(* IEC 61131-3 sources: JingjiangArm/moonboxpro_arm_8.4/Application/Application/任务列表/ExtTask/动作处理/涂布, 11 files *)

(* ---- StCoatingAxisInf.st ---- *)
(*@CES
Name=StCoatingAxisInf
Type=Gvl
TypeGuid=2db5746d-d284-4425-9f7f-2663a34b0ebc
Guid=2e9ecafb-d2f1-4b6b-83e3-f47895db637f
HasDeclaration=True
HasImplementation=False
*)
{DECLARATION}
TYPE StCoatingAxisInf :
STRUCT
(*涂布轴信息@2024.01.18.095207*)
	byCoatingAxisNum			: BYTE;(*涂布轴个数*)
	aiAxisIdList				: ARRAY [1..gc_byCoatingMaxSum_New]OF INT;(*轴idlist*)
	astStCoatingAxisParam		: ARRAY [1..gc_byCoatingMaxSum_New] OF StCoatingAxisParam;
END_STRUCT
END_TYPE

{IMPLEMENTATION}

(* ---- StCoatingAxisParam.st ---- *)
(*@CES
Name=StCoatingAxisParam
Type=Gvl
TypeGuid=2db5746d-d284-4425-9f7f-2663a34b0ebc
Guid=8a071cba-fd95-4a8c-93c6-fe3e9b0305b5
HasDeclaration=True
HasImplementation=False
*)
{DECLARATION}
{attribute 'pack_mode' := '1'}
TYPE StCoatingAxisParam :(*涂布轴参数@2024.01.18.093551*)
STRUCT
	iUnitId							:INT;(*轴id@默认-1*)
	xSwitchOn_CoatingPrn			:BOOL;(*涂布开关*)
	byAdjMode_CoatingPrn			:BYTE;(*涂布轴模式*)
	xReverseAdj_CoatingPrn			:BOOL;(*涂布轴调整取反*)
	rAI_CoatingPrn					:REAL;(*涂布轴模拟量*)
	rAI_med_CoatingPrn				:REAL;(*涂布轴中位值*)
	lrGirth_Using_CoatingPrn		:LREAL;(*涂布轴周长@界面输入*)
	iKp_CoatingPrn					:INT;(*涂布kp*)
	iKi_CoatingPrn					:INT;(*涂布ki*)
	iKd_CoatingPrn					:INT;(*涂布kd*)
	xFlag_PressDne					:BOOL;(*涂布轴合压*)

	rAI_CoatingHMI					:REAL;(*涂布模拟量显示*)
	lrGirth_CoatingPrn				:LREAL;(*涂布周长@用于运算pt*)
	lrVelocity_CoatingPrn			:LREAL;(*涂布速度*)
END_STRUCT
END_TYPE

{IMPLEMENTATION}

(* ---- KS_CoatingAxisParamDeal.st ---- *)
(*@CES
Name=KS_CoatingAxisParamDeal
Type=FunctionBlock
TypeGuid=6f9dac99-8de1-4efc-8465-68ac443b7d08
Guid=f4156371-7451-43fd-b965-d24d4d478a2f
HasDeclaration=True
HasImplementation=True
*)
{DECLARATION}
FUNCTION KS_CoatingAxisParamDeal : BOOL
VAR_INPUT
(*涂布轴参数处理*)
	i_byDealType:BYTE;(*处理方式@=1 初始化涂布轴参数
								@=2 从轴参数写入到涂布轴参数中#涂布控制输入变量
								@=3 涂布轴参数写入到轴参数中#涂布控制输出变量
								@=4 操作的轴参数值复位*)
	i_iAxisId:INT;
	i_xFlag_AxisPressDne:BOOL;(*轴的合压状态@经过延时后输出标志*)
	i_pstStCoatingAxisParam:POINTER TO StCoatingAxisParam;
	i_palrGirth_CoatingPrn:POINTER TO ARRAY [1..MAX_UNIT_NUM] OF LREAL;(*用于计算pt的周长值@未定义到轴参数中*)
	i_palrAI_CoatingHMI:POINTER TO ARRAY [1..MAX_UNIT_NUM] OF LREAL;(*界面显示的模拟量值@未定义到轴参数中*)
//2025.7.3.175755
	i_axSwitchOn_CoatingPrn: ARRAY [1..MAX_UNIT_NUM] OF BOOL;(*涂布开关*)
	i_abyAdjMode_CoatingPrn: ARRAY [1..MAX_UNIT_NUM] OF BYTE;(*涂布轴模式*)
	i_axReverseAdj_CoatingPrn: ARRAY [1..MAX_UNIT_NUM] OF BOOL;(*涂布轴调整取反*)
	i_alrAI_CoatingPrn: ARRAY [1..MAX_UNIT_NUM] OF LREAL;(*涂布模拟量*)
	i_alrAI_med_CoatingPrn: ARRAY [1..MAX_UNIT_NUM] OF LREAL;(*涂布中位值*)
	i_alrGirth_Using_CoatingPrn: ARRAY [1..MAX_UNIT_NUM] OF LREAL;(*涂布轴周长*)
	i_aiKp_CoatingPrn: ARRAY [1..MAX_UNIT_NUM] OF INT;(*涂布Kp*)
	i_aiKi_CoatingPrn: ARRAY [1..MAX_UNIT_NUM] OF INT;(*涂布Ki*)
	i_aiKd_CoatingPrn: ARRAY [1..MAX_UNIT_NUM] OF INT;(*涂布Kd*)
	i_palrVelocity_CoatingPrn:POINTER TO ARRAY [1..MAX_UNIT_NUM] OF LREAL;(*涂布轴速度*)
	i_alrGirth:ARRAY [1..MAX_UNIT_NUM] OF LREAL;(*当前轴周长*)
END_VAR
VAR
END_VAR

{IMPLEMENTATION}
CASE i_byDealType OF
	1:(*初始化涂布参数*)
		IF i_pstStCoatingAxisParam<>0 THEN
			SysMemSet(i_pstStCoatingAxisParam,0,SIZEOF(i_pstStCoatingAxisParam^));
			i_pstStCoatingAxisParam^.iUnitId:=-1;
		END_IF
	2:(*从轴参数写入到涂布轴参数中#涂布控制输入变量*)
		IF i_iAxisId>0 AND i_iAxisId<MAX_UNIT_NUM AND(*轴号合法*)

			i_pstStCoatingAxisParam<>0 THEN

			i_pstStCoatingAxisParam^.iUnitId						:= i_iAxisId;
			i_pstStCoatingAxisParam^.xSwitchOn_CoatingPrn			:= i_axSwitchOn_CoatingPrn[i_iAxisId];(*涂布开关*)
			i_pstStCoatingAxisParam^.byAdjMode_CoatingPrn			:= i_abyAdjMode_CoatingPrn[i_iAxisId];(*涂布轴模式*)
			i_pstStCoatingAxisParam^.xReverseAdj_CoatingPrn			:= i_axReverseAdj_CoatingPrn[i_iAxisId]	;(*涂布轴调整取反*)
			i_pstStCoatingAxisParam^.rAI_CoatingPrn					:= i_alrAI_CoatingPrn[i_iAxisId];(*涂布轴模拟量*)
			i_pstStCoatingAxisParam^.rAI_med_CoatingPrn				:= i_alrAI_med_CoatingPrn[i_iAxisId];(*涂布轴中位值*)
			i_pstStCoatingAxisParam^.lrGirth_Using_CoatingPrn		:= i_alrGirth_Using_CoatingPrn[i_iAxisId];(*涂布轴周长@界面输入*)
			i_pstStCoatingAxisParam^.iKp_CoatingPrn					:= i_aiKp_CoatingPrn[i_iAxisId]	;(*涂布kp*)
			i_pstStCoatingAxisParam^.iKi_CoatingPrn					:= i_aiKi_CoatingPrn[i_iAxisId];(*涂布ki*)
			i_pstStCoatingAxisParam^.iKd_CoatingPrn					:= i_aiKd_CoatingPrn[i_iAxisId]	;(*涂布kd*)
			i_pstStCoatingAxisParam^.xFlag_PressDne					:= i_xFlag_AxisPressDne			;(*涂布轴合压*)
		END_IF
	3:(*涂布轴参数写入到轴参数中*)
		IF i_iAxisId>0 AND i_iAxisId<MAX_UNIT_NUM AND(*轴号合法*)
			i_pstStCoatingAxisParam<>0 AND
			i_palrGirth_CoatingPrn<>0 AND
			i_palrAI_CoatingHMI<>0 THEN

			i_palrAI_CoatingHMI^[i_iAxisId]			:= i_pstStCoatingAxisParam^.rAI_CoatingHMI		 	;(*涂布模拟量显示*)
			i_palrGirth_CoatingPrn^[i_iAxisId]		:= i_pstStCoatingAxisParam^.lrGirth_CoatingPrn	 	;(*涂布周长@用于运算pt*)
			i_palrVelocity_CoatingPrn^[i_iAxisId]	:= i_pstStCoatingAxisParam^.lrVelocity_CoatingPrn	;(*涂布速度*)
		END_IF

	4:(*操作的轴参数值复位*)
		IF i_iAxisId>0 AND i_iAxisId<MAX_UNIT_NUM AND(*轴号合法*)
			i_palrGirth_CoatingPrn<>0 AND
			i_palrAI_CoatingHMI<>0 THEN

			i_palrAI_CoatingHMI^[i_iAxisId]			:= 0;(*涂布模拟量显示*)
			i_palrGirth_CoatingPrn^[i_iAxisId]		:= i_alrGirth[i_iAxisId];(*赋值为当前周长*)
			i_palrVelocity_CoatingPrn^[i_iAxisId]	:= 0;(*涂布速度*)
		END_IF
ELSE;(*啥也不干*)
END_CASE

(* ---- KS_GetCoatingAllnf.st ---- *)
(*@CES
Name=KS_GetCoatingAllnf
Type=FunctionBlock
TypeGuid=6f9dac99-8de1-4efc-8465-68ac443b7d08
Guid=cb71e24b-1db6-4b3f-8052-350591e92417
HasDeclaration=True
HasImplementation=True
*)
{DECLARATION}
FUNCTION KS_GetCoatingAllnf : bool
(*获取系轴中涂布模拟量@未做滤波(如果需要可以在获取的地方进行运算)*)
VAR_INPUT
	i_xGetCoatingAxisAI:BOOL;(*获取涂布轴ai*)
	i_xGetUnitAxisAI:BOOL;(*获取所有色组轴ai*)
	i_rPressure_Max:REAL;(*压力传感器最大值*)
	i_iGrpAxisNum_Pu: INT;(*色组轴数量|*)
	i_paiGrpAxisList: POINTER TO ARRAY [1..MAX_UNIT_NUM] OF INT;(*系轴列表|有排序规则|*)
	i_pstStCoatingAxisInf:POINTER TO StCoatingAxisInf;
	i_pastStIOMap_AxisExtra:POINTER TO ARRAY [1..MAX_UNIT_NUM] OF StIOMap_Axis_Extra_FE;
	i_paiAIAxisIdlist_Last:POINTER TO ARRAY[1..MAX_UNIT_NUM] OF INT;(*获取ai的轴id列表备份*)
	i_pabySensorType_CoatingPrn:POINTER TO ARRAY[1..MAX_UNIT_NUM] OF BYTE;(*涂布传感器类型*)
	i_abyAdjMode_CoatingPrn:ARRAY[1..MAX_UNIT_NUM] OF BYTE;
	i_palrAI_CoatingPrn:POINTER TO ARRAY [1..MAX_UNIT_NUM] OF LREAL;
END_VAR
VAR
	iN: INT;
	iM: INT;
	iNum: INT:=0;
	aiIdlist: ARRAY [1..MAX_UNIT_NUM] OF INT:=[(-1)];
	iUnitId: INT;
	pstStIOMap_AxisExtra:POINTER TO StIOMap_Axis_Extra_FE;
	iTemp: INT;
	lrMinTemp: LREAL;
	lrMaxTemp: LREAL;
	diMinTemp: DINT;
	diMaxTemp: DINT;
	lrTemp: LREAL;
END_VAR
{IMPLEMENTATION}
IF i_pstStCoatingAxisInf<>0 AND
	i_paiGrpAxisList<>0 AND
	i_pastStIOMap_AxisExtra<>0 AND
	i_paiAIAxisIdlist_Last<>0 THEN;
ELSE
	RETURN;
END_IF

IF i_xGetCoatingAxisAI THEN(*获取涂布轴ai*)
	iNum:=i_pstStCoatingAxisInf^.byCoatingAxisNum;
	FOR iN:=1 TO i_pstStCoatingAxisInf^.byCoatingAxisNum BY 1 DO
		aiIdlist[iN]:=i_pstStCoatingAxisInf^.aiAxisIdList[iN];
	END_FOR
ELSIF i_xGetUnitAxisAI THEN(*获取所有色组轴ai*)
	iNum:=i_iGrpAxisNum_Pu;
	FOR iN:=1 TO i_pstStCoatingAxisInf^.byCoatingAxisNum BY 1 DO
		aiIdlist[iN]:=i_paiGrpAxisList^[iN];
	END_FOR
ELSE;
END_IF

FOR iN:=1 TO iNum BY 1 DO
	iUnitId:=aiIdlist[iN];
	IF iUnitId>0 AND iUnitId<=MAX_UNIT_NUM THEN
		pstStIOMap_AxisExtra:=ADR(i_pastStIOMap_AxisExtra^[iUnitId]);

		(*获取配置的类型*)
		i_pabySensorType_CoatingPrn^[iUnitId]:=0;
		IF pstStIOMap_AxisExtra^.i_byAIType_CoatingSensor<=5 THEN
			i_pabySensorType_CoatingPrn^[iUnitId]:=pstStIOMap_AxisExtra^.i_byAIType_CoatingSensor;
		END_IF

		(*获取配置的模拟值@转换未正负*)
		iTemp:=WORD_TO_INT(pstStIOMap_AxisExtra^.i_wAI_CoatingSensor);

		(*获取上下限*)
		KS_QueryRangeByAType(
							i_pabySensorType_CoatingPrn^[iUnitId],
							ADR(lrMinTemp),
							ADR(lrMaxTemp),
							ADR(diMinTemp),
							ADR(diMaxTemp));

		(*计算模拟量值*)
		i_palrAI_CoatingPrn^[iUnitId]:=KSIO_DA(iTemp,
												lrMinTemp,
												lrMaxTemp,
												diMinTemp,
												diMaxTemp);

		(*增加了张力传感器时的显示值处理2019.8.9.161738*)
		IF lrMinTemp<0 THEN lrMinTemp:=0;END_IF(*最小值是负值的传感器一般0--正模拟量值对应0--最大量*)
		lrTemp:=lrMaxTemp-lrMinTemp;
		IF lrTemp<>0 THEN;ELSE lrTemp:=10;END_IF(*按照0--10v处理*)

		IF i_abyAdjMode_CoatingPrn[iUnitId]=2 OR i_abyAdjMode_CoatingPrn[iUnitId]=3 THEN
		(*张力传感器调整时，将电压值转换为张力值*)
			lrTemp:=i_rPressure_Max(*pstStGrpParam^.rPressure_Max*)/lrTemp;(*默认最小压力为0*)
			i_palrAI_CoatingPrn^[iUnitId]:=(i_palrAI_CoatingPrn^[iUnitId]-lrMinTemp)*lrTemp;
		END_IF
	END_IF
END_FOR

(*寻找消失的轴*)
FOR iN:=1 TO MAX_UNIT_NUM BY 1 DO
	iUnitId:=i_paiAIAxisIdlist_Last^[iN];(*之前的轴id*)
	IF iUnitId>0 AND iUnitId<=MAX_UNIT_NUM  THEN
		IF iNum>0 THEN
			FOR iM:=1 TO iNum BY 1 DO
				IF aiIdlist[iM]=iUnitId THEN(*还在呢*)
					EXIT;
				ELSE(*已经被删除了*)
					IF iM=iNum THEN(*列表里没了*)
						i_palrAI_CoatingPrn^[iUnitId]:=0;(*复位操作的值*)
					END_IF
				END_IF
			END_FOR
		ELSE(*一个都没有 就把之前的关闭把*)
			//pstStAxisParam:=ADR(i_pastStAxisParam^[iUnitId]);
			i_palrAI_CoatingPrn^[iUnitId]:=0;(*复位操作的值*)
		END_IF
	END_IF
END_FOR

i_paiAIAxisIdlist_Last^:=aiIdlist;(*备份列表值*)

(* ---- KS_GetCoatingAxisInf.st ---- *)
(*@CES
Name=KS_GetCoatingAxisInf
Type=FunctionBlock
TypeGuid=6f9dac99-8de1-4efc-8465-68ac443b7d08
Guid=94653cdc-8513-44b1-a378-a0e4607a5782
HasDeclaration=True
HasImplementation=True
*)
{DECLARATION}
FUNCTION KS_GetCoatingAxisInf : BOOL
VAR_INPUT
(*获取涂布轴参数@2024.01.18.094943*)
	i_pstStCoatingAxisInf:POINTER TO StCoatingAxisInf;
	i_paxFlag_PressDne:POINTER TO ARRAY [1..MAX_UNIT_NUM] OF BOOL;
	i_palrGirth_CoatingPrn:POINTER TO ARRAY [1..MAX_UNIT_NUM] OF LREAL;(*用于计算pt的周长值@未定义到轴参数中*)
	//2025.07.22.105010
	i_axSwitchOn_CoatingPrn: ARRAY [1..MAX_UNIT_NUM] OF BOOL;(*涂布开关*)
	i_abyAdjMode_CoatingPrn: ARRAY [1..MAX_UNIT_NUM] OF BYTE;(*涂布轴模式*)
	i_axReverseAdj_CoatingPrn: ARRAY [1..MAX_UNIT_NUM] OF BOOL;(*涂布轴调整取反*)
	i_alrAI_CoatingPrn: ARRAY [1..MAX_UNIT_NUM] OF LREAL;(*涂布模拟量*)
	i_alrAI_med_CoatingPrn: ARRAY [1..MAX_UNIT_NUM] OF LREAL;(*涂布中位值*)
	i_alrGirth_Using_CoatingPrn: ARRAY [1..MAX_UNIT_NUM] OF LREAL;(*涂布轴周长*)
	i_aiKp_CoatingPrn: ARRAY [1..MAX_UNIT_NUM] OF INT;(*涂布Kp*)
	i_aiKi_CoatingPrn: ARRAY [1..MAX_UNIT_NUM] OF INT;(*涂布Ki*)
	i_aiKd_CoatingPrn: ARRAY [1..MAX_UNIT_NUM] OF INT;(*涂布Kd*)
	i_palrVelocity_CoatingPrn:POINTER TO ARRAY [1..MAX_UNIT_NUM] OF LREAL;(*涂布轴速度*)
	i_alrGirth:ARRAY [1..MAX_UNIT_NUM] OF LREAL;(*当前轴周长*)
END_VAR
VAR
	iN: INT;
	iUnitId: INT;
	xFlag_AxisPressDne: BOOL;
	byDealType: BYTE;(*处理方式@=1 初始化涂布轴参数
								@=2 从轴参数写入到涂布轴参数中#涂布控制输入变量
								@=3 涂布轴参数写入到轴参数中#涂布控制输出变量
								@=4 操作的轴参数值复位*)
END_VAR

{IMPLEMENTATION}
IF i_pstStCoatingAxisInf<>0 AND
	i_paxFlag_PressDne<>0 AND
	i_palrGirth_CoatingPrn<>0 THEN;
ELSE
	RETURN;
END_IF

(*初始化和获取涂布轴参数*)
FOR iN:=1 TO gc_byCoatingMaxSum_New BY 1 DO
	iUnitId:=i_pstStCoatingAxisInf^.aiAxisIdList[iN];(*之前的轴id*)
	IF iUnitId=-1 THEN(*无效则清除参数*)
		byDealType:=1;
	ELSE(*ID有效@加载参数*)
		byDealType:=2;
		xFlag_AxisPressDne:=i_paxFlag_PressDne^[iUnitId];(*获取新轴的参数*)
	END_IF
	KS_CoatingAxisParamDeal(
		byDealType(*i_byDealType*) ,
		iUnitId(*i_iAxisId*) ,
		xFlag_AxisPressDne(*i_xFlag_AxisPressDne*) ,
		ADR(i_pstStCoatingAxisInf^.astStCoatingAxisParam[iN])(*i_pstStCoatingAxisParam*) ,
		i_palrGirth_CoatingPrn(*i_palrGirth_CoatingPrn*) ,
		0(*i_palrAI_CoatingHMI*) ,
		i_axSwitchOn_CoatingPrn(*i_axSwitchOn_CoatingPrn*) ,
		i_abyAdjMode_CoatingPrn(*i_abyAdjMode_CoatingPrn*),
		i_axReverseAdj_CoatingPrn(*i_axReverseAdj_CoatingPrn*),
		i_alrAI_CoatingPrn(*i_alrAI_CoatingPrn*),
		i_alrAI_med_CoatingPrn(*i_alrAI_med_CoatingPrn*),
		i_alrGirth_Using_CoatingPrn(*i_alrGirth_Using_CoatingPrn*),
		i_aiKp_CoatingPrn(*i_aiKp_CoatingPrn*),
		i_aiKi_CoatingPrn(*i_aiKi_CoatingPrn*),
		i_aiKd_CoatingPrn(*i_aiKd_CoatingPrn*),
		i_palrVelocity_CoatingPrn(*i_palrVelocity_CoatingPrn*),
		i_alrGirth(*i_alrGirth*) );

END_FOR

(* ---- KS_GetCoatingAxisList.st ---- *)
(*@CES
Name=KS_GetCoatingAxisList
Type=FunctionBlock
TypeGuid=6f9dac99-8de1-4efc-8465-68ac443b7d08
Guid=8bc67aac-0c7f-4420-a195-db7a2a94b6c1
HasDeclaration=True
HasImplementation=True
*)
{DECLARATION}
FUNCTION KS_GetCoatingAxisList : BOOL
VAR_INPUT
	i_iGrpAxisNum_Pu: INT;(*色组轴数量|*)
	i_paiGrpAxisList: POINTER TO ARRAY [1..MAX_UNIT_NUM] OF INT;(*系轴列表|有排序规则|*)
	i_pstStCoatingAxisInf:POINTER TO StCoatingAxisInf;
	i_axSwitchOn_CoatingPrn: ARRAY [1..MAX_UNIT_NUM] OF BOOL;
END_VAR
VAR
	iN: INT;
	iUnitId: INT;
	aiAxisIdList:ARRAY [1..gc_byCoatingMaxSum_New] OF INT;(*2024.01.18.104002*)
	byCoatingNum: BYTE;
END_VAR

{IMPLEMENTATION}
IF i_pstStCoatingAxisInf<>0 AND
	i_paiGrpAxisList<>0THEN;
ELSE
	RETURN;
END_IF

(*处理涂布轴列表*)
byCoatingNum:=0;
FOR iN:=1 TO gc_byCoatingMaxSum_New BY 1 DO
	aiAxisIdList[iN]:=-1;
END_FOR

FOR iN:=1 TO i_iGrpAxisNum_Pu BY 1 DO
	iUnitId:=i_paiGrpAxisList^[iN];
	IF iUnitId>0 AND iUnitId<=MAX_UNIT_NUM THEN
		IF i_axSwitchOn_CoatingPrn[iUnitId] THEN(*涂布打开*)
			byCoatingNum:=byCoatingNum+1;
			IF byCoatingNum<=gc_byCoatingMaxSum_New THEN(*不能超过可以处理的个数*)
				aiAxisIdList[byCoatingNum]:=iUnitId;
				IF byCoatingNum=gc_byCoatingMaxSum_New THEN
					EXIT;
				END_IF
			END_IF
		END_IF
	END_IF
END_FOR
(*写入到结构体中*)
i_pstStCoatingAxisInf^.byCoatingAxisNum:=byCoatingNum;
i_pstStCoatingAxisInf^.aiAxisIdList:=aiAxisIdList;

(* ---- KS_SetCoatingAxisInf.st ---- *)
(*@CES
Name=KS_SetCoatingAxisInf
Type=FunctionBlock
TypeGuid=6f9dac99-8de1-4efc-8465-68ac443b7d08
Guid=aab75e54-4a14-456c-b5e5-3fbc7559278d
HasDeclaration=True
HasImplementation=True
*)
{DECLARATION}
FUNCTION KS_SetCoatingAxisInf : bool
(*设置涂布轴信息@写入到轴参数中*)
VAR_INPUT
	i_pstStCoatingAxisInf:POINTER TO StCoatingAxisInf;
	i_aiAxisIdList_Last:POINTER TO ARRAY [1..gc_byCoatingMaxSum_New]OF INT;(*备份的轴列表*)
	i_palrGirth_CoatingPrn:POINTER TO ARRAY [1..MAX_UNIT_NUM] OF LREAL;(*用于计算pt的周长值@未定义到轴参数中*)
	i_palrAI_CoatingHMI:POINTER TO ARRAY [1..MAX_UNIT_NUM] OF LREAL;(*界面显示的模拟量值@未定义到轴参数中*)
		//2025.07.22.105010
	i_axSwitchOn_CoatingPrn: ARRAY [1..MAX_UNIT_NUM] OF BOOL;(*涂布开关*)
	i_abyAdjMode_CoatingPrn: ARRAY [1..MAX_UNIT_NUM] OF BYTE;(*涂布轴模式*)
	i_axReverseAdj_CoatingPrn: ARRAY [1..MAX_UNIT_NUM] OF BOOL;(*涂布轴调整取反*)
	i_alrAI_CoatingPrn: ARRAY [1..MAX_UNIT_NUM] OF LREAL;(*涂布模拟量*)
	i_alrAI_med_CoatingPrn: ARRAY [1..MAX_UNIT_NUM] OF LREAL;(*涂布中位值*)
	i_alrGirth_Using_CoatingPrn: ARRAY [1..MAX_UNIT_NUM] OF LREAL;(*涂布轴周长*)
	i_aiKp_CoatingPrn: ARRAY [1..MAX_UNIT_NUM] OF INT;(*涂布Kp*)
	i_aiKi_CoatingPrn: ARRAY [1..MAX_UNIT_NUM] OF INT;(*涂布Ki*)
	i_aiKd_CoatingPrn: ARRAY [1..MAX_UNIT_NUM] OF INT;(*涂布Kd*)
	i_palrVelocity_CoatingPrn:POINTER TO ARRAY [1..MAX_UNIT_NUM] OF LREAL;(*涂布轴速度*)
	i_alrGirth:ARRAY [1..MAX_UNIT_NUM] OF LREAL;(*当前轴周长*)
END_VAR
VAR
	iN: INT;
	iM: INT;
	iUnitId: INT;
	byDealType: BYTE;(*处理方式@=1 初始化涂布轴参数
								@=2 从轴参数写入到涂布轴参数中#涂布控制输入变量
								@=3 涂布轴参数写入到轴参数中#涂布控制输出变量
								@=4 操作的轴参数值复位*)
	aiAxisIdList_Last:ARRAY [1..gc_byCoatingMaxSum_New] OF INT;(*2024.01.18.104002*)
END_VAR

{IMPLEMENTATION}
IF i_pstStCoatingAxisInf<>0 AND
	i_aiAxisIdList_Last<>0 AND
	i_palrGirth_CoatingPrn<>0 AND
	i_palrAI_CoatingHMI<>0 THEN;
ELSE
	RETURN;
END_IF
aiAxisIdList_Last:=i_aiAxisIdList_Last^;(*获取*)

(*设置涂布轴参数*)
FOR iN:=1 TO i_pstStCoatingAxisInf^.byCoatingAxisNum BY 1 DO
	iUnitId:=i_pstStCoatingAxisInf^.aiAxisIdList[iN];(*现在轴id*)
	IF iUnitId=-1 THEN(*无效则*)
		byDealType:=0;(*啥也不干*)
	ELSE(*ID有效@写入到轴参数中*)
		byDealType:=3;
	END_IF

	KS_CoatingAxisParamDeal(
		byDealType(*i_byDealType*) ,
		iUnitId(*i_iAxisId*) ,
		FALSE(*i_xFlag_AxisPressDne*) ,
		ADR(i_pstStCoatingAxisInf^.astStCoatingAxisParam[iN])(*i_pstStCoatingAxisParam*) ,
		i_palrGirth_CoatingPrn(*i_palrGirth_CoatingPrn*) ,
		i_palrAI_CoatingHMI(*i_palrAI_CoatingHMI*) ,
		i_axSwitchOn_CoatingPrn(*i_axSwitchOn_CoatingPrn*) ,
		i_abyAdjMode_CoatingPrn(*i_abyAdjMode_CoatingPrn*),
		i_axReverseAdj_CoatingPrn(*i_axReverseAdj_CoatingPrn*),
		i_alrAI_CoatingPrn(*i_alrAI_CoatingPrn*),
		i_alrAI_med_CoatingPrn(*i_alrAI_med_CoatingPrn*),
		i_alrGirth_Using_CoatingPrn(*i_alrGirth_Using_CoatingPrn*),
		i_aiKp_CoatingPrn(*i_aiKp_CoatingPrn*),
		i_aiKi_CoatingPrn(*i_aiKi_CoatingPrn*),
		i_aiKd_CoatingPrn(*i_aiKd_CoatingPrn*),
		i_palrVelocity_CoatingPrn(*i_palrVelocity_CoatingPrn*),
		i_alrGirth(*i_alrGirth*) );
END_FOR

FOR iN:=1 TO gc_byCoatingMaxSum_New BY 1 DO
	iUnitId:=aiAxisIdList_Last[iN];(*之前的轴id*)
	IF iUnitId>0 AND iUnitId<=MAX_UNIT_NUM THEN
		byDealType:=0;
		IF i_pstStCoatingAxisInf^.byCoatingAxisNum>0 THEN
			FOR iM:=1 TO i_pstStCoatingAxisInf^.byCoatingAxisNum BY 1 DO
				IF i_pstStCoatingAxisInf^.aiAxisIdList[iM]=iUnitId THEN(*还在呢*)
					EXIT;
				ELSE(*已经被删除了*)
					IF iM=i_pstStCoatingAxisInf^.byCoatingAxisNum THEN(*列表里没了*)
						byDealType:=4;(*复位操作的值*)
					END_IF
				END_IF
			END_FOR
		ELSE(*一个都没有*)
			byDealType:=4;(*复位操作的值*)
		END_IF

	KS_CoatingAxisParamDeal(
		byDealType(*i_byDealType*) ,
		iUnitId(*i_iAxisId*) ,
		FALSE(*i_xFlag_AxisPressDne*) ,
		ADR(i_pstStCoatingAxisInf^.astStCoatingAxisParam[iN])(*i_pstStCoatingAxisParam*) ,
		i_palrGirth_CoatingPrn(*i_palrGirth_CoatingPrn*) ,
		i_palrAI_CoatingHMI(*i_palrAI_CoatingHMI*) ,
		i_axSwitchOn_CoatingPrn(*i_axSwitchOn_CoatingPrn*) ,
		i_abyAdjMode_CoatingPrn(*i_abyAdjMode_CoatingPrn*),
		i_axReverseAdj_CoatingPrn(*i_axReverseAdj_CoatingPrn*),
		i_alrAI_CoatingPrn(*i_alrAI_CoatingPrn*),
		i_alrAI_med_CoatingPrn(*i_alrAI_med_CoatingPrn*),
		i_alrGirth_Using_CoatingPrn(*i_alrGirth_Using_CoatingPrn*),
		i_aiKp_CoatingPrn(*i_aiKp_CoatingPrn*),
		i_aiKi_CoatingPrn(*i_aiKi_CoatingPrn*),
		i_aiKd_CoatingPrn(*i_aiKd_CoatingPrn*),
		i_palrVelocity_CoatingPrn(*i_palrVelocity_CoatingPrn*),
		i_alrGirth(*i_alrGirth*) );
	END_IF
END_FOR

aiAxisIdList_Last:=i_pstStCoatingAxisInf^.aiAxisIdList;(*更新备份的涂布轴列表*)
i_aiAxisIdList_Last^:=aiAxisIdList_Last;(*写入*)

(* ---- KS_FB_CalGirthByVel.st ---- *)
(*@CES
Name=KS_FB_CalGirthByVel
Type=FunctionBlock
TypeGuid=6f9dac99-8de1-4efc-8465-68ac443b7d08
Guid=9f5d0384-92e8-4505-b8ed-e463be3a3529
HasDeclaration=True
HasImplementation=True
*)
{DECLARATION}
FUNCTION_BLOCK KS_FB_CalGirthByVel
VAR_INPUT
	i_xEn:BOOL;(**)
	i_iCycleTime:INT;(*程序执行周期*)
	i_lrAnalog: LREAL;(*模拟量输入相对于中位差值变量*)
	i_rAnalogLimit:REAL;(*模拟量的限值*)
	i_lrFilmVel:LREAL;(*料膜速度值*)
	i_lrVel:LREAL;(*当前周期的调整速度值*)
	i_lrUsingGirth:LREAL;(*使用的周长值*)
	i_rAnalogSumLimit:REAL;(*模拟量累计值的限值*)
END_VAR
VAR_OUTPUT
	o_xEn:BOOL;
	o_xGirthCaled:BOOL;(*周长计算完成了~*)
	o_lrGirth:LREAL;(*计算出来的周长值*)
END_VAR
VAR

	iCycleCount: INT:=0;(*周期计数值*)
	lrCurrentVelSum:LREAL;(*当前速度累计值*)
	iN: INT;
	lrAnalogSum: LREAL;(*当前模拟量的累计值*)
	lrAver_CurrentVel: LREAL;

	alrDataFifo:ARRAY [1..2,1..c_iArrNum] OF LREAL;(*用来存放每个周期速度以及模拟量的值。一维数组代表速度值，二维数组代表模拟量值*)
	xArrInited: BOOL;(*数组初始完成*)
	iLastIndex: INT;(*100个周期之前的模拟量数据索引*)
	xAnalogValue: BOOL;(*模拟量有效*)
	iDelayCount: INT;
END_VAR
VAR CONSTANT
	c_iArrNum:INT:=100;(*数组大小暂定为100个 按20ms周期算就是2s的数据*)
END_VAR

{IMPLEMENTATION}
o_xGirthCaled:=FALSE;(*该标志只有效一个周期*)
o_lrGirth:=0;
lrAver_CurrentVel:=0;
lrCurrentVelSum:=0;
lrAnalogSum:=0;
IF i_xEn  THEN(*使能计算周长功能*)

(*保存一定时间的速度值，用来进行平均速度计算。时间暂定为2s*)
	iCycleCount:=iCycleCount+1;(*计数+1*)
	IF iCycleCount>c_iArrNum THEN(*循环存储*)
		iCycleCount:=1;
	END_IF
	alrDataFifo[1,iCycleCount]:=i_lrVel;(*速度值*)
	alrDataFifo[2,iCycleCount]:=i_lrAnalog;(*模拟量值*)

	IF iCycleCount>=c_iArrNum OR xArrInited THEN (*累计足够次数的速度值*)
		xArrInited:=TRUE;
		iDelayCount:=iDelayCount+1;
	(*计算模拟量累计值和速度累计值*)
		FOR iN:=1 TO c_iArrNum BY 1 DO
			lrCurrentVelSum:=lrCurrentVelSum+alrDataFifo[1,iN];
			IF ABS(alrDataFifo[2,iN])>i_rAnalogLimit AND iDelayCount<=500 THEN
				(*2020.3.5.104548_|iDelayCount<=300修改到500|*)
					(*累计的这段时间里的模拟量值必须都小于等于模拟量限值才有效
											iDelayCount 是用来保证在极端情况下不能满足条件也可以进入计算逻辑*)
				lrAnalogSum:=i_rAnalogSumLimit+1;(*给模拟量累计值一个大于模拟量累计限值的值，这样我们在下面的判断中则会认为无效*)
				xAnalogValue:=FALSE;
				EXIT;
			ELSE
				xAnalogValue:=TRUE;
				lrAnalogSum:=lrAnalogSum+alrDataFifo[2,iN];
			END_IF
		END_FOR

(*修改计算平均速度的条件2018.5.8.121744*)
(*(*原条件*)
		IF ABS(lrAnalogSum)>i_rAnalogSumLimit THEN(*模拟量累计值超过范围，则认为无效*);
		ELSE(*模拟量累计值在一定范围内求取速度平均值*)
			lrAver_CurrentVel:=lrCurrentVelSum/INT_TO_LREAL(c_iArrNum);
		END_IF
*)
		iLastIndex:=(iCycleCount+1) MOD c_iArrNum;

		IF (ABS((alrDataFifo[2,iCycleCount])-(alrDataFifo[2,iLastIndex])) >0.005) OR (NOT  xAnalogValue) THEN(*模拟量2S的变化量超过范围，则认为无效*);
		ELSE(*模拟量累计值在一定范围内求取速度平均值*)
			lrAver_CurrentVel:=lrCurrentVelSum/INT_TO_LREAL(c_iArrNum);
		END_IF
	END_IF

	IF lrAver_CurrentVel<>0 AND i_lrFilmVel<>0 THEN (*平均速度不等于0 我们认为已经计算出了满足条件的平均速度值*)
		o_lrGirth:=i_lrFilmVel*i_lrUsingGirth/lrAver_CurrentVel;(*计算出理论周长值*)
		o_xGirthCaled:=TRUE;
	END_IF

ELSE
	iDelayCount:=0;
	iCycleCount:=0;
	xArrInited:=FALSE;
END_IF
o_xEn:=i_xEn;

(* ---- KS_FB_CalGirthLogic_Coating.st ---- *)
(*@CES
Name=KS_FB_CalGirthLogic_Coating
Type=FunctionBlock
TypeGuid=6f9dac99-8de1-4efc-8465-68ac443b7d08
Guid=e8f75550-8c47-4eed-8c0f-4881fe2307b6
HasDeclaration=True
HasImplementation=True
*)
{DECLARATION}
FUNCTION_BLOCK KS_FB_CalGirthLogic_Coating
VAR_INPUT
	i_xEn:BOOL;
	i_xAdjNewWay:BOOL;(*调整算法新方法使能标志，在计算完成后直接进行周长自增自减调整*)
	i_xGirthAdj:BOOL;(*新算法中周长调整使能*)(*2019.8.9.155755修改为直接启动周长自增自减标志*)
	i_xCompensate_Dir:BOOL;
	(*模拟量输入和中位差值与料膜松紧关系标志：FALSE： 差值大于0代表料松，小于0代表料紧、TRUE ：差值大于0代表料紧，小于0代表料松*)
	i_iCycleTime:INT;(*程序执行周期*)
	i_lrAnalog:LREAL;(*模拟量值，摆臂位置*)
	i_rAnalogLimit:REAL;(*模拟量有效值限值*)
	i_lrFilmVel:LREAL;(*料膜速度*)
	i_lrVel:LREAL;(*实际速度*)
	i_lrActualGirth:LREAL;(*默认周长*)
END_VAR
VAR_OUTPUT
	o_xEn:BOOL;
	o_xGirthCalFinish:BOOL;(*计算完成标志有效了 就不在进行调整*)
	o_lrUsingGirth:LREAL;
END_VAR
VAR
	fbKS_FB_CalGirthByVel: KS_FB_CalGirthByVel;
	xGirthCaled: BOOL;
	lrGirthTemp: LREAL;
	xCalGirthEn: BOOL;(*计算周长使能标志*)
	xEvenning: BOOL;(*匀速标志*)
	lrPreCurVel: LREAL;
	xPreGirthCalFinish: BOOL;
	xInit: BOOL;

	lrAnalog_Aver: LREAL:=0;
	lrPreAnalog_Aver: LREAL;
(*	rGirthStep:REAL:=0.01;(*周长变化步进量*)*)
	rGirthStep:REAL:=0.02; (* 2020.7.13.094914|重现调整数值 *)

	lrAnalog_Sum: LREAL;
	xCalAverDone: BOOL;
	rThreshold: REAL;
	iCycleCount:INT;
	iCoeff: INT;
	iCalGirthCount: INT;
	xConditionDone: BOOL;
	lrGirthStep_Temp: LREAL;
	iThreshold: INT:=5;(*计算出的的牵引周长有效范围单位%*)
END_VAR
VAR CONSTANT
	(*2020.4.22.101241|新增|*)
	c_lrAIBoundage_Axis: LREAL := 0.8;
END_VAR

{IMPLEMENTATION}
(*稳速时候才能进行周长计算*)
xEvenning:=FALSE;
IF i_lrFilmVel=lrPreCurVel AND i_lrFilmVel>=10  THEN(*速度大于一定值，并且处于匀速*)
	xEvenning:=TRUE;
END_IF

xConditionDone:=FALSE;
IF xEvenning THEN(*进入匀速状态之后 等待一段时间在进入计算周长状态*)
	iCalGirthCount:=iCalGirthCount+1;
	IF iCalGirthCount>=500 THEN (*延迟500个周期 进入计算周长状态*)
		iCalGirthCount:=iCalGirthCount-1;
		xConditionDone:=TRUE;
	END_IF
ELSE
	iCalGirthCount:=0;
END_IF

xCalGirthEn:=FALSE;
IF xConditionDone AND (NOT o_xGirthCalFinish) AND i_xAdjNewWay(*g_xInFeedAndOutFeed_AdjNewWay *)THEN
	xCalGirthEn:=TRUE;
END_IF

fbKS_FB_CalGirthByVel(
	i_xEn:=xCalGirthEn ,
	i_iCycleTime:=i_iCycleTime ,
	i_lrAnalog:=i_lrAnalog ,
	i_rAnalogLimit:=i_rAnalogLimit ,
	i_lrFilmVel:=i_lrFilmVel ,
	i_lrVel:=i_lrVel ,
	i_lrUsingGirth:= o_lrUsingGirth,
	i_rAnalogSumLimit:=,
	o_xEn=> ,
	o_xGirthCaled=> xGirthCaled,
	o_lrGirth=>lrGirthTemp );

IF xGirthCaled THEN
	o_xGirthCalFinish:=TRUE;(*该标志有效则可以认为我们可以进入非调整状态了*)
END_IF

IF o_xGirthCalFinish AND ABS(i_lrAnalog)>c_lrAIBoundage_Axis THEN(*2020.4.22.101215_|0.3--->>>c_lrAIBoundage_Axis|*)
	o_xGirthCalFinish:=FALSE;
END_IF

IF o_xGirthCalFinish AND (NOT xPreGirthCalFinish)  THEN(*将计算出来的值赋给输出值*)
	IF lrGirthTemp<=i_lrActualGirth*(1+iThreshold/100.0) AND lrGirthTemp>=i_lrActualGirth*(1-iThreshold/100.0) THEN
		o_lrUsingGirth:=lrGirthTemp;
	ELSE
		o_xGirthCalFinish:=FALSE;
	END_IF
END_IF

IF   i_lrFilmVel=0 THEN(*不走料的时候版周长为默认值*)
	(*IF   NOT xInit THEN*)
		o_xGirthCalFinish:=FALSE;
		o_lrUsingGirth:=i_lrActualGirth;
		xInit:=TRUE;
(*	END_IF*)
ELSE
	xInit:=FALSE;
END_IF

(*当已经进入到不再调整逻辑中的时候，我们对牵引的周长进行微调*)(*2018.5.7.153458*)

(*求摆臂的位置的平均值*)
xCalAverDone:=FALSE;
iCycleCount:=iCycleCount+1;
lrAnalog_Sum:=lrAnalog_Sum+i_lrAnalog;
IF iCycleCount>=50 THEN
	xCalAverDone:=TRUE;
	(*lrPreAnalog_Aver:=lrAnalog_Aver;*)
	lrAnalog_Aver:=lrAnalog_Sum/iCycleCount;
	lrAnalog_Sum:=0;
	iCycleCount:=0;
ELSE;
END_IF

IF o_xGirthCalFinish AND (NOT xPreGirthCalFinish)  THEN(*计算完成后初始化上个周期平均模拟量值*)
	lrPreAnalog_Aver:=lrAnalog_Aver;
END_IF

lrGirthTemp:=0;
lrGirthStep_Temp:=rGirthStep;
IF (o_xGirthCalFinish OR i_xGirthAdj(*g_xGirthAdj  *)) AND xCalAverDone THEN
	IF ABS(lrAnalog_Aver)>0.1 THEN
		rThreshold:=0;
	ELSE
		rThreshold:=0.001;
	END_IF

	IF NOT  i_xCompensate_Dir THEN(*对于补偿方向取反*)
		iCoeff:=1;
	ELSE
		iCoeff:=-1;
	END_IF

	IF  lrAnalog_Aver >0.01 THEN
		IF  lrAnalog_Aver>lrPreAnalog_Aver+rThreshold THEN(*位置值越来越大了*)
			lrGirthTemp:=iCoeff*lrGirthStep_Temp;
			lrPreAnalog_Aver:=lrAnalog_Aver;
		END_IF
	ELSIF  lrAnalog_Aver <-0.01  THEN
		IF  lrAnalog_Aver+rThreshold<lrPreAnalog_Aver THEN(*位置值越来越小了*)
			lrGirthTemp:=-iCoeff*lrGirthStep_Temp;
			lrPreAnalog_Aver:=lrAnalog_Aver;
		END_IF
	ELSE
		lrPreAnalog_Aver:=lrAnalog_Aver;
	END_IF
ELSE;
END_IF

o_lrUsingGirth:=o_lrUsingGirth+lrGirthTemp;

lrPreCurVel:=i_lrFilmVel;
xPreGirthCalFinish:=o_xGirthCalFinish;
o_xEn:=i_xEn;

(* ---- KS_FB_Coating_Tension.st ---- *)
(*@CES
Name=KS_FB_Coating_Tension
Type=FunctionBlock
TypeGuid=6f9dac99-8de1-4efc-8465-68ac443b7d08
Guid=b2750bde-e2fb-4c3e-bf55-6bf4b42d8bc9
HasDeclaration=True
HasImplementation=True
*)
{DECLARATION}
FUNCTION_BLOCK KS_FB_Coating_Tension(*涂布张力算法|传感器有两种：1是使用PI调整计算周长调整周长；2是使用周长调整*)
(*张力调整方式:
0-手动调整周长
1-摆臂调整方式下,稳定后调整周长
2-张力传感器方式下,稳定后调整周长
3-张力传感器下直接调整周长
4-摆臂方式下,一直使用pid(2022.10.24.205316)*)
(*调整速度限值值修改到2--10m/min*)
VAR_INPUT
	i_xEn:BOOL;(*涂布张力使能*)
	i_xCoatingAdjDir:BOOL;(*涂布调整方向*)
	i_byCoatingAdjWay:BYTE;(*调整方式:0为不自动调整；1为摆臂模式*)
	i_lrCurrentVel:LREAL;(*当前速度*)
	i_lrFilmVel:LREAL;(*料膜速度*)
	i_lrCoatingGirth:LREAL;(*涂布版周长*)
	i_lrAnalog:LREAL;(*相对于中位的模拟量值*)
	i_lrP:LREAL;
	i_lrD:LREAL;
	(*pi限制值单位%|2022.10.13.124543*)
	i_byVelLimit_PerCent:BYTE;(*速度限制百分比%*)
END_VAR
VAR_OUTPUT
	o_xEn:BOOL;(**)
	o_lrCoatingVel:LREAL;(*涂布速度*)
	o_lrCoatingUsingGirth:LREAL;(*涂布使用的版周长*)
END_VAR
VAR

	alrArrDataBak			: ARRAY [1..10] OF LREAL;

	lrCoatingPI_Value		: LREAL;
	iCoeff					: INT;
	rMaxDelVel				: REAL;(*单个周期最大的调整量*)
	lrAddValue				: LREAL:=0;(*叠加的调整量*)
	iVelocityLimit			: INT:=10;(*速度限值 *)
	xCoatingPIAdj			: BOOL:=FALSE;
	fbKS_FB_CalGirthLogic	: KS_FB_CalGirthLogic_Coating;(*周长调整功能块*)
	iN						: INT;
	xCoatAdjFlag			: BOOL;(*涂布调整标志*)

	xGirthCalFinish			: BOOL;
	lrDel					: LREAL:=0;
	iDataBak_Index: INT;
END_VAR

{IMPLEMENTATION}
(*根据调整速度计算版周长 并进行补偿*)
fbKS_FB_CalGirthLogic(
	i_xEn:=TRUE,
	i_xAdjNewWay:=i_xEn AND (i_byCoatingAdjWay=1 OR i_byCoatingAdjWay=2) ,
						(*进行摆臂涂布调整或者张力传感器1的时候 才进行周长的计算以及补偿*)
	i_xGirthAdj:=i_xEn AND (i_byCoatingAdjWay=3),(*张力传感器2的方式直接调整版周长*)
	i_xCompensate_Dir:= (NOT i_xCoatingAdjDir),
	i_iCycleTime:=gc_TENSION_TSK_CYCLE_TIME ,
	i_lrAnalog:=i_lrAnalog ,
	i_rAnalogLimit:=0.1,
	i_lrFilmVel:=i_lrFilmVel ,
	i_lrVel:=o_lrCoatingVel,
	i_lrActualGirth:=i_lrCoatingGirth ,
	o_xEn=> ,
	o_xGirthCalFinish=>xGirthCalFinish,
	o_lrUsingGirth=>o_lrCoatingUsingGirth );

xCoatingPIAdj:=i_byCoatingAdjWay=4 OR(*2022.10.24.205601 增加了摆臂方式下pi常调整方式*)
			((i_byCoatingAdjWay=1 OR i_byCoatingAdjWay=2) AND NOT xGirthCalFinish);(*摆臂调整时 并且周长未计算完成则进行调整*)

(*涂布调整手动调整会保存在周长值中。若是自动调整的周长值则不会保存*)
IF i_byCoatingAdjWay=0 OR (*涂布周长手动调整*)
	i_byCoatingAdjWay=4 THEN(*2022.10.24.205710 增加*)
	o_lrCoatingUsingGirth:=i_lrCoatingGirth;
ELSIF i_byCoatingAdjWay=1 OR i_byCoatingAdjWay=2(*涂布摆臂调整或者)*)
		OR i_byCoatingAdjWay=3 THEN(*张力传感器方式1时*);
END_IF

o_xEn:=i_xEn;
rMaxDelVel:=0.3;(*=300/20/50 20S加速到300m/min的时候一个周期速度的变化量*)(*2018.5.22.115216 增加调整量限值*)

(*2022.10.13.124549 速度限制使用%|最小2m/min 最大10m/min*)
IF i_byVelLimit_PerCent<>0 THEN
	iVelocityLimit:=LREAL_TO_INT(i_byVelLimit_PerCent*i_lrFilmVel/100);
ELSE(*等于0按照10m/min限制-以前一直使用该值*)
	iVelocityLimit:=10;
END_IF

IF iVelocityLimit<2 THEN
	iVelocityLimit:=2;
ELSIF iVelocityLimit>10 THEN
	iVelocityLimit:=10;
END_IF

IF i_lrFilmVel=0 THEN(*料膜速度为0速的时候，调整牵引到中位。对速度进行限值*)(*2018.7.11.223054*)
	iVelocityLimit:=2;
END_IF

FOR iN:=10 TO 2 BY -1 DO
	alrArrDataBak[iN]:=alrArrDataBak[iN-1];
END_FOR
alrArrDataBak[1]:=i_lrAnalog;

IF i_xEn THEN(*涂布调整使能*)
	(*2020.5.11.163738 尝试将pd值的输入值
	相比以前放大10倍。并将d值的差值改为和上个周期的。*)
	iDataBak_Index:=5;
	IF i_byCoatingAdjWay=2 THEN
		i_lrP:=i_lrP/100;
		i_lrD:=i_lrD/100;
		iDataBak_Index:=2;
	END_IF

	lrCoatingPI_Value:=i_lrP/1000*(i_lrAnalog)+
						i_lrD/100*(alrArrDataBak[1]-alrArrDataBak[iDataBak_Index]);

	iCoeff:=1;
	IF i_xCoatingAdjDir THEN iCoeff:=-1; END_IF(*控制pi调整方向*)

	lrCoatingPI_Value:=lrCoatingPI_Value*iCoeff;

	IF i_byCoatingAdjWay=0 OR i_byCoatingAdjWay=3 THEN(*若为手动调整或者张力传感器方式2。不改变速度*)
		lrCoatingPI_Value:=0;
	END_IF

	IF ABS(lrCoatingPI_Value)>rMaxDelVel THEN(*对调整量进行限值*)
		lrCoatingPI_Value:=rMaxDelVel*lrCoatingPI_Value/ABS(lrCoatingPI_Value);
	END_IF

	lrAddValue:=lrAddValue+lrCoatingPI_Value;
	IF ABS(lrAddValue)>iVelocityLimit THEN
		lrAddValue:=iVelocityLimit*ABS(lrAddValue)/lrAddValue;
	END_IF

	o_lrCoatingVel:=i_lrCurrentVel+lrAddValue;

	IF xCoatingPIAdj THEN(*涂布速度pi调整*);
	ELSE(*不再速度pi调整，使用调整周长的方式*)
		IF i_byCoatingAdjWay=1 OR i_byCoatingAdjWay=2 THEN
			o_lrCoatingVel:=i_lrCurrentVel;
			lrAddValue:=0;
		END_IF
	END_IF
	xCoatAdjFlag:=TRUE;
	lrDel:=(lrAddValue)/1000;(*1s减速到0*)
ELSE(**)
	IF i_lrCurrentVel=0 THEN
		IF xCoatAdjFlag THEN xCoatAdjFlag:=FALSE; END_IF
	END_IF

	IF lrAddValue>0 THEN
		lrAddValue:=lrAddValue-lrDel*gc_TENSION_TSK_CYCLE_TIME;
		IF lrAddValue <0 THEN
			lrAddValue:=0;
		END_IF
	ELSIF lrAddValue<0 THEN
		lrAddValue:=lrAddValue-lrDel*gc_TENSION_TSK_CYCLE_TIME;
		IF lrAddValue >0 THEN
			lrAddValue:=0;
		END_IF
	ELSE
		lrDel:=0;
	END_IF
	o_lrCoatingVel:=i_lrCurrentVel+lrAddValue;
END_IF

IF o_lrCoatingVel<0 THEN o_lrCoatingVel:=0;END_IF

(* ---- KS_FB_CoatingCTL.st ---- *)
(*@CES
Name=KS_FB_CoatingCTL
Type=FunctionBlock
TypeGuid=6f9dac99-8de1-4efc-8465-68ac443b7d08
Guid=407fa95c-6cd2-4404-bcf4-68a89e2fd197
HasDeclaration=True
HasImplementation=True
*)
{DECLARATION}
FUNCTION_BLOCK KS_FB_CoatingCTL
VAR_INPUT
	i_xEn: BOOL;
	i_iGrpId: INT;
	i_iGrpAxisNum_Pu: INT;(*色组轴数*)
	i_aiGrpAxisList: ARRAY [1..MAX_UNIT_NUM] OF INT;(*系轴列表*)
	i_pastStIOMap_AxisBasic:POINTER TO ARRAY [1..MAX_UNIT_NUM] OF StIOMap_Main_FE;
	i_pastStIOMap_AxisExtra:POINTER TO ARRAY [1..MAX_UNIT_NUM] OF StIOMap_Axis_Extra_FE;
	i_pstStCoatingAxisInf:POINTER TO StCoatingAxisInf;
	i_pstStSysParam: POINTER TO StSysParam;
	i_paxFlag_PressDne:POINTER TO ARRAY [1..MAX_UNIT_NUM] OF BOOL;
	i_palrGirth_CoatingPrn:POINTER TO ARRAY [1..MAX_UNIT_NUM] OF LREAL;(*用于计算pt的周长值@未定义到轴参数中*)
	i_palrAI_CoatingHMI:POINTER TO ARRAY [1..MAX_UNIT_NUM] OF LREAL;(*界面显示的模拟量值@未定义到轴参数中*)
END_VAR
VAR_OUTPUT
END_VAR
VAR
	iN: INT;
	iUnitId: INT;
//	iGrp:INT;
	//iCoatId:INT;
	lrTemp: LREAL;
	iMaxTemp: INT;
	lrAIDel: LREAL;
	xNotCoatingUnitPressed: BOOL;
	xFlag_PressDne: BOOL;
	afbKS_FB_Coating_Tension: ARRAY [1.. gc_byCoatingMaxSum_New] OF KS_FB_Coating_Tension;
	aiAxisIdList_Last:ARRAY [1..gc_byCoatingMaxSum_New] OF INT;(*2024.01.18.104002*)
	xTensionCtlEn: BOOL;
	iIndex: INT;

//2026.8.20.170304	lrGirth_Using_CoatingPrn_In:ARRAY[1..MAX_UNIT_NUM] OF LREAL;(*使用的涂布版周长*)
	xLinkage_In:ARRAY[1..MAX_UNIT_NUM] OF BOOL;(*轴联动状态*)
	rVel_Film_In: REAL;(*料膜速度*)
	byVelLimit_PerCent_IfOf_In: BYTE;(*速度限制百分比*)
	rVel_Cur_In: REAL;(*当前速度*)
	axSwitchOn_CoatingPrn_In: ARRAY [1..MAX_UNIT_NUM] OF BOOL;
	abyAdjMode_CoatingPrn_In: ARRAY [1..MAX_UNIT_NUM] OF BYTE;(*涂布轴模式*)
	axReverseAdj_CoatingPrn_In: ARRAY [1..MAX_UNIT_NUM] OF BOOL;(*涂布轴调整取反*)
	alrAI_CoatingPrn_In: ARRAY [1..MAX_UNIT_NUM] OF LREAL;(*涂布模拟量*)
	alrAI_med_CoatingPrn_In: ARRAY [1..MAX_UNIT_NUM] OF LREAL;(*涂布中位值*)
	alrGirth_Using_CoatingPrn_In: ARRAY [1..MAX_UNIT_NUM] OF LREAL;(*涂布轴周长*)
	aiKp_CoatingPrn_In: ARRAY [1..MAX_UNIT_NUM] OF INT;(*涂布Kp*)
	aiKi_CoatingPrn_In: ARRAY [1..MAX_UNIT_NUM] OF INT;(*涂布Ki*)
	aiKd_CoatingPrn_In: ARRAY [1..MAX_UNIT_NUM] OF INT;(*涂布Kd*)
	alrVelocity_CoatingPrn_In: ARRAY [1..MAX_UNIT_NUM] OF LREAL;(*涂布速度*)
	alrGirth_In:ARRAY[1..MAX_UNIT_NUM] OF LREAL;(*当前轴周长*)
	rPressure_Max_In:LREAL;(*压力传感器最大值*)
	aiAIAxisIdlist_Last_In:ARRAY[1..MAX_UNIT_NUM] OF INT;(*获取ai的轴id列表备份*)
	abySensorType_CoatingPrn_In: ARRAY [1..MAX_UNIT_NUM] OF BYTE;(*传感器类型*)
	byCoatingAxisNum_In:BYTE;(*涂布轴个数*)
//	aiAxisIdList_In:ARRAY[1..gc_byCoatingMaxSum_New] OF INT;(*涂布轴列表*)
//	xSwitchOn_CoatingPrn_In:ARRAY[1..gc_byCoatingMaxSum_New] OF BOOL;(*涂布开关*)
//	byAdjMode_CoatingPrn_In:ARRAY[1..gc_byCoatingMaxSum_New] OF BYTE;(*涂布轴模式*)
//	xReverseAdj_CoatingPrn_In:ARRAY[1..gc_byCoatingMaxSum_New] OF BOOL;(*涂布轴调整取反*)
//	rAI_CoatingPrn_In:ARRAY[1..gc_byCoatingMaxSum_New] OF REAL;(*涂布轴模拟量*)
//	rAI_med_CoatingPrn_In:ARRAY[1..gc_byCoatingMaxSum_New] OF REAL;(*涂布轴中位值*)
//	lrGirth_Using_CoatingPrnHMI_In:ARRAY[1..gc_byCoatingMaxSum_New] OF LREAL;(*涂布轴周长@界面输入*)
//	iKp_CoatingPrn_In:ARRAY[1..gc_byCoatingMaxSum_New] OF INT;(*涂布kp*)
//	iKi_CoatingPrn_In:ARRAY[1..gc_byCoatingMaxSum_New] OF INT;(*涂布ki*)
//	iKd_CoatingPrn_In:ARRAY[1..gc_byCoatingMaxSum_New] OF INT;(*涂布kd*)
//	xFlag_PressDne_In:ARRAY[1..gc_byCoatingMaxSum_New] OF BOOL;(*涂布轴合压*)
//	rAI_CoatingHMI_In:ARRAY[1..gc_byCoatingMaxSum_New] OF REAL;(*涂布模拟量显示*)
//	lrGirth_CoatingPrn_In:ARRAY[1..gc_byCoatingMaxSum_New] OF LREAL;(*涂布周长@用于运算pt*)
//	lrVelocity_CoatingPrn_In:ARRAY[1..gc_byCoatingMaxSum_New] OF LREAL;(*涂布速度*)

	abyAxisList_CoatingPrn_Out:ARRAY[1..MAX_UNIT_NUM] OF BYTE;(*涂布轴列表*)
	byAxisNum_CoatingPrn_Out:BYTE;(*涂布轴个数*)
	pstStCoatingAxisParam:POINTER TO StCoatingAxisParam;
//	aiAxisIdList_Last:ARRAY [1..gc_byCoatingMaxSum_New] OF INT;(*2024.01.18.104002*)
END_VAR

{IMPLEMENTATION}
Action_Input();
Action_Act();
Action_Output();
